// TIA Portal V20 export
FUNCTION_BLOCK "FB_VFD"   // FB103, LAD
TITLE = Variable speed drive with speed monitoring
{ S7_Optimized_Access := 'TRUE' }
AUTHOR : Demo
VERSION : 0.2
// LAD version. Same interface as scl/15_FB_VFD.scl.
// stored: AutoNumber false, SetENOAutomatically false
   VAR_INPUT
      Run : Bool;   // Request: run the drive
      Permit : Bool := true;   // Interlock: drive may only run when TRUE
      SpeedSP : Real;   // Requested speed [rpm]
      SpeedPV : Real;   // Actual speed from the drive [rpm]
      Ready : Bool;   // Drive ready
      DriveFault : Bool;   // Drive reports a fault
      DeviationTime : Time := T#15S;   // How long speed may be too low before a fault
   END_VAR
   VAR_OUTPUT
      RunOut : Bool;   // Run command to the drive
      SpeedOut : Real;   // Speed setpoint to the drive [rpm]
      AtSpeed : Bool;   // Actual speed within 10 % of setpoint
      FaultDrive : Bool;   // Drive fault
      FaultSpeedDev : Bool;   // Running, but speed more than 10 % below setpoint for DeviationTime
      NotReady : Bool;   // Drive not ready (and no fault): check enable / E-stop / main switch
   END_VAR
   VAR
      tDev : TON_TIME;   // Speed deviation time
   END_VAR
   VAR_TEMP
      SpeedMin : Real;   // 90 % of the speed setpoint [rpm]
   END_VAR
BEGIN

REGION Network 1: Drive fault
   // The drive reports a fault.
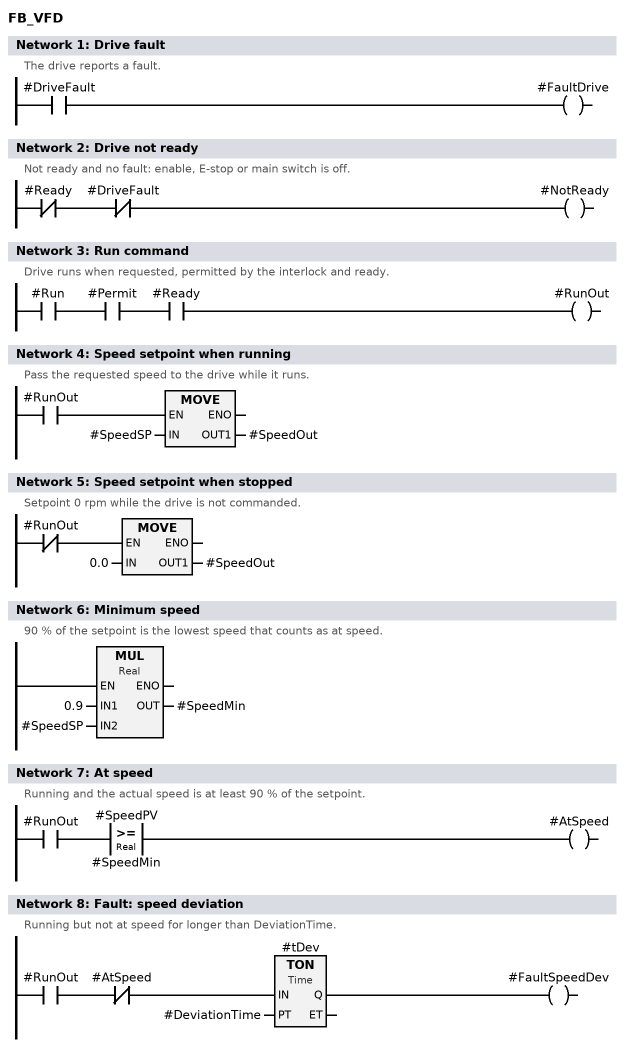
   RUNG wire#powerrail
      Contact( #DriveFault )
      Coil( #FaultDrive )
   END_RUNG
   // the same network as SCL:
   #FaultDrive := #DriveFault;
END_REGION

REGION Network 2: Drive not ready
   // Not ready and no fault: enable, E-stop or main switch is off.
   RUNG wire#powerrail
      I_Contact( #Ready )
      I_Contact( #DriveFault )
      Coil( #NotReady )
   END_RUNG
   // the same network as SCL:
   #NotReady := NOT #Ready AND NOT #DriveFault;
END_REGION

REGION Network 3: Run command
   // Drive runs when requested, permitted by the interlock and ready.
   RUNG wire#powerrail
      Contact( #Run )
      Contact( #Permit )
      Contact( #Ready )
      Coil( #RunOut )
   END_RUNG
   // the same network as SCL:
   #RunOut := #Run AND #Permit AND #Ready;
END_REGION

REGION Network 4: Speed setpoint when running
   // Pass the requested speed to the drive while it runs.
   RUNG wire#powerrail
      Contact( #RunOut )
      { S7_GenerateENO := "TRUE" } Move(in := #SpeedSP, out1 => #SpeedOut)
   END_RUNG
   // the same network as SCL:
   IF #RunOut THEN #SpeedOut := #SpeedSP; END_IF;
END_REGION

REGION Network 5: Speed setpoint when stopped
   // Setpoint 0 rpm while the drive is not commanded.
   RUNG wire#powerrail
      I_Contact( #RunOut )
      { S7_GenerateENO := "TRUE" } Move(in := 0.0, out1 => #SpeedOut)
   END_RUNG
   // the same network as SCL:
   IF NOT #RunOut THEN #SpeedOut := 0.0; END_IF;
END_REGION

REGION Network 6: Minimum speed
   // 90 % of the setpoint is the lowest speed that counts as at speed.
   RUNG wire#powerrail
      { S7_Templates := "SrcType := Real"; S7_GenerateENO := "TRUE" } Mul(in1 := 0.9, in2 := #SpeedSP, out => #SpeedMin)
   END_RUNG
   // the same network as SCL:
   #SpeedMin := 0.9 * #SpeedSP;
END_REGION

REGION Network 7: At speed
   // Running and the actual speed is at least 90 % of the setpoint.
   RUNG wire#powerrail
      Contact( #RunOut )
      { S7_Templates := "SrcType := Real" } GE_Contact(in1 := #SpeedPV, in2 := #SpeedMin)
      Coil( #AtSpeed )
   END_RUNG
   // the same network as SCL:
   #AtSpeed := #RunOut AND (#SpeedPV >= #SpeedMin);
END_REGION

REGION Network 8: Fault: speed deviation
   // Running but not at speed for longer than DeviationTime.
   RUNG wire#powerrail
      Contact( #RunOut )
      I_Contact( #AtSpeed )
      { S7_Templates := "time_type := Time" } #tDev.TON(pt := #DeviationTime, et =>)
      Coil( #FaultSpeedDev )
   END_RUNG
   // the same network as SCL:
   #tDev(IN := #RunOut AND NOT #AtSpeed, PT := #DeviationTime);   // TON
   #FaultSpeedDev := #tDev.Q;
END_REGION
END_FUNCTION_BLOCK
